FUNCTION_BLOCK EV_NeedleAxis (* Names the equipment's two channels, and unpacks its state channel into named values (its inputs and who holds it) for a skill. Technical: Names NeedleAxis's channels; typed view of its state channel (inputs and holder) *)
  (* Standard: 61499-2 *)
  (* Version 0.1, 2026-09-28, Project contributors, AAU Smart Production Lab *)
  PACKAGE filler;
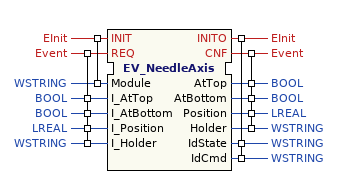
  EVENT_INPUT
    INIT : EInit WITH Module; (* Name the equipment's channels *)
    REQ WITH I_AtTop, I_AtBottom, I_Position, I_Holder; (* The equipment's state arrived *)
  END_EVENT
  EVENT_OUTPUT
    INITO : EInit WITH IdState, IdCmd; (* IdState and IdCmd are set *)
    CNF WITH AtTop, AtBottom, Position, Holder; (* The values below are updated *)
  END_EVENT
  VAR_INPUT
    Module : WSTRING; (* The module's name; its local channels are named after it (loc[<Module>/...]) *)
    I_AtTop : BOOL; (* AtTop as read or received *)
    I_AtBottom : BOOL; (* AtBottom as read or received *)
    I_Position : LREAL; (* Position as read or received *)
    I_Holder : WSTRING; (* Holder as read or received *)
  END_VAR
  VAR_OUTPUT
    AtTop : BOOL; (* NeedleAxis: AtTop, an input *)
    AtBottom : BOOL; (* NeedleAxis: AtBottom, an input *)
    Position : LREAL; (* NeedleAxis: Position (mm), an input *)
    Holder : WSTRING; (* Who holds the equipment (empty: free) *)
    IdState : WSTRING; (* Local channel of the equipment's state *)
    IdCmd : WSTRING; (* Local channel of the equipment's commands *)
  END_VAR
  EC_STATES
    INIT : INIT -> INITO;
    REQ : REQ -> CNF;
  END_STATES
  ALGORITHM INIT IN ST:
IdState := CONCAT(CONCAT("loc[", Module), "/NeedleAxis/state]");
IdCmd := CONCAT(CONCAT("loc[", Module), "/NeedleAxis/cmd]");
  END_ALGORITHM
  ALGORITHM REQ IN ST:
AtTop := I_AtTop;
AtBottom := I_AtBottom;
Position := I_Position;
Holder := I_Holder;
  END_ALGORITHM
END_FUNCTION_BLOCK
